// TIA Portal V20 export
// export: Created 2026-10-19T18:45:26.87382Z, ExportSetting None, DisplayName Totally Integrated Automation Portal, DisplayVersion V20 Update 6, DisplayName TIA Portal Openness, DisplayVersion V20 Update 6, DisplayName TIA Portal Version Control Interface, DisplayVersion V20 Update 6, DisplayName SINAMICS Startdrive Advanced, DisplayVersion V20 SP1, DisplayName SINAMICS Startdrive G130, G150, S120, S150, SINAMICS MV, G220, S200, S210, DisplayVersion V20 SP1, DisplayName SINAMICS Startdrive G110M, G120, G120C, G120D, G120P, G115D, DisplayVersion V20 SP1, DisplayName STEP 7 Professional, DisplayVersion V20 Update 6, DisplayName STEP 7 Safety, DisplayVersion V20 Update 2, DisplayName WinCC Basic/Comfort/Advanced, DisplayVersion V20 Update 6, DisplayName WinCC Unified, DisplayVersion V20 Update 6
VAR_GLOBAL   // PLC tag table "IO_ET200_1"
   "VTD1 LEVEL DETECT 1" AT %I10.0 : Bool;
   "VTD1 LEVEL DETECT 2" AT %I10.1 : Bool;
   "C1103 STOPPER RAISED" AT %I5.0 : Bool;
   "C1103 STOPPER LOWERED" AT %I5.1 : Bool;
   "C1103 STOPPER MOTOR" AT %Q5.4 : Bool;
   "C1104 STOPPER MOTOR" AT %Q6.4 : Bool;
   "C1104 STOPPER RAISED" AT %I6.0 : Bool;
   "C1104 STOPPER LOWERED" AT %I6.1 : Bool;
   "C1106 STOPPER RAISED" AT %I8.0 : Bool;
   "C1105 STOPPER RAISED" AT %I7.0 : Bool;
   "C1105 STOPPER MOTOR" AT %Q7.4 : Bool;
   "C1105 STOPPER LOWERED" AT %I7.1 : Bool;
   "C1106 STOPPER MOTOR" AT %Q8.4 : Bool;
   "C1102 STOPPER MOTOR" AT %Q4.4 : Bool;
   "C1106 STOPPER LOWERED" AT %I8.1 : Bool;
   "C1102 STOPPER LOWERED" AT %I4.1 : Bool;
   "VTD1 DOCKING PINS RETRACTED 2" AT %I9.2 : Bool;
   "OVERTRAVEL LOWER LIMIT - CH2(1)" AT %I528.4 : Bool;
   "C1102 STOPPER RAISED" AT %I4.0 : Bool;
   "VTD1 DOCKING PINS RETRACTED 1" AT %I9.3 : Bool;
   "OVERTRAVEL UPPER LIMIT - CH1(1)" AT %I528.1 : Bool;
   "VTD1 DOCKING PINS 1 EXTEND" AT %Q9.4 : Bool;
   "VTD1 DOCKING PINS EXTENDED 2" AT %I9.1 : Bool;
   "VTD1 DOCKING PINS 2 EXTEND" AT %Q9.5 : Bool;
   "VTD1 DOCKING PINS EXTENDED 1" AT %I9.0 : Bool;
   "VTD1 DOCKING PINS 1 RETRACT" AT %Q9.6 : Bool;
   "OVERTRAVEL LOWER LIMIT - CH1(1)" AT %I528.0 : Bool;
   "OVERTRAVEL UPPER LIMIT - CH2(1)" AT %I528.5 : Bool;
   "VTD1 DOCKING PINS 2 RETRACT" AT %Q9.7 : Bool;
END_VAR
